PROGRAM PRG_Main
VAR
    fbMachine : FB_IndexedPatchPressMachine;
END_VAR

fbMachine.Cyclic(
    stInputs := GVL_MASTER.stInputs,
    stCommand := GVL_MASTER.stCommand,
    stConfig := GVL_Config.stMachine,
    bPatchDispenseCommissioned := GVL_PatchPress_Interface.bPatchDispenseCommissioned,
    bHeatStakeCommissioned := GVL_PatchPress_Interface.bHeatStakeCommissioned,
    bVisionCommissioned := GVL_PatchPress_Interface.bVisionCommissioned,
    bCoreCommissioningMode := GVL_PatchPress_Interface.bCoreCommissioningMode,
    bLogoutHMI := FALSE,
    stOutputs => GVL_MASTER.stOutputs,
    stStatus => GVL_MASTER.stStatus);

END_PROGRAM

(* stored: Version 1.1.0.1, ProductVersion 3.1.4026.18
   POU PRG_Main: Id {fe8f5db4-2dbe-44c9-ba3e-79c06469fde0}, SpecialFunc None *)
